Fanuc KAREL source: kd00059.KL

-- PROVISIONAL review KL for V770-1; original PC SHA256 d87a2bc2c7e4bc11b5fe0761d5d4a1b9c7341eec384e2b152efc1e4eee8e6d22
-- Incomplete behavior may be omitted. Consult companion uncertainty JSON. Do not deploy.
PROGRAM KD00059
%NOLOCKGROUP
VAR
  I : INTEGER
  J : INTEGER
  B : BOOLEAN
  R : REAL
  S : STRING[80]
BEGIN
  -- UNRESOLVED_PC offsets 5-18; opcodes 9D,81,18,9D,1B,9D,12,9C,13,04
  -- UNRESOLVED_PC offsets 23-27; opcodes 7F
END KD00059
